Fanuc KAREL source: KB00053.KL

PROGRAM KB00053
%NOLOCKGROUP
%ENVIRONMENT BYNAM
VAR
  RESULT: STRING[80]
BEGIN
  RESULT = CURR_PROG
END KB00053
